TYPE ST_Prod_Ingredient :
STRUCT
	sDescription		: STRING:= 'Ingredient Name';
	eIngredientType		: E_Ingredient_type;
	rWeight				: REAL; // kg
	rWeightPercentage	: REAL;
	rFlowRate_Dissolving: REAL;
	rFlowRate_Blending	: REAL;
	tBlendingDuration	: TIME;

END_STRUCT
END_TYPE

(* stored: Version 1.1.0.1, ProductVersion 3.1.4024.15
   DUT ST_Prod_Ingredient: Id {a004cfa8-fe17-41ed-9ff5-bd508f086eec} *)
